Fanuc KAREL source: kd00049.KL

-- PROVISIONAL review KL for V770-1; original PC SHA256 f265c7c56201906678ab7a94682f42b8419948620c3153a303ed2be49112ebb9
-- Incomplete behavior may be omitted. Consult companion uncertainty JSON. Do not deploy.
PROGRAM KD00049
%NOLOCKGROUP
VAR
  I : INTEGER
  J : INTEGER
  B : BOOLEAN
  R : REAL
  S : STRING[80]
BEGIN
  -- UNRESOLVED_PC offsets 5-18; opcodes 01,2E,0A,82,0B
  -- UNRESOLVED_PC offsets 23-27; opcodes 7F
END KD00049
